(* IEC 61131-3 sources: SortJet_MasterSPS_Aufbau.fbsproj/09_Station/Stationen/_Basic, 3 files *)

(* ---- Basic_Glastransport_FB_V01_00_00.fb.st ---- *)
(* METADATA
{
	"v3Meta": {
		"objectGuid": "8cc859a4-3853-4716-ad69-f1a04cff8809"
	}
}
*)
FUNCTION_BLOCK Basic_Glastransport_FB_V01_00_00
VAR_INPUT

  // BOOL
  bpAktivieren                     : BOOL;
  bpEintransport                   : BOOL;
  bpEintransportRueckwaertig       : BOOL;
  bpAustransport                   : BOOL;
  bpAustransportRueckwaertig       : BOOL;
  bpVortransport                   : BOOL;
  bpVortransportRueckwaertig       : BOOL;
  bpMesskopplung                   : BOOL;
  bpDurchtransport                 : BOOL;
  bpGlaslaengenmessung             : BOOL;
  bpHandfahrenPlus                 : BOOL;
  bpHandfahrenMinus                : BOOL;
  bpScheibeZurueckFahren           : BOOL;
  bpScheibeVorFahren               : BOOL;
  bpAnforderungHandfunktion        : BOOL; // Handfunktionen greifen auch im Automatikbetrieb (z.B. waehrend der Bediener anlegt)
  bpScheibeQuittiert               : BOOL; // Bediener hat die Scheibe quittiert (Fehlmessung / Messergebnis)
  bpScheibeFreigegeben             : BOOL; // Scheibe ist nach der Messung freigegeben
  bpReferenz                       : BOOL;
  bpCheck                          : BOOL;
  bpReset                          : BOOL;
  bpAutomatikAktiv                 : BOOL;
  bpFreigabe                       : BOOL;
  bpMessrichtungNegativ            : BOOL;
  bpCheckMitVorgaenger             : BOOL;
  bpCheckMitNachfolger             : BOOL;
  bpRueckwaertigerTransport        : BOOL;
  bpScheibentrennen                : BOOL;
  bpAbbruchVortransport            : BOOL;

  // Sensoren
  bpSensorEinlauf                  : BOOL;
  bpSensorEinlaufVorAb             : BOOL;
  bpSensorAuslaufVorAb             : BOOL;
  bpSensorAuslauf                  : BOOL;

  // OPTIONEN
  bpOptionMessungSystemCheckAktiv            : BOOL;
  bpOptionMasterSlaveTransport               : BOOL;
  bpOptionScheibenmessungEintransport        : BOOL;
  bpOptionAustransportISOLinie               : BOOL;
  bpOptionSlaveAntrieb                       : BOOL;
  bpOptionNachSystemcheckAufAuslaufsensor    : BOOL;
  bpOptionbScheibenmessungSensorVorabAuslauf : BOOL;

  // WORD
  wlIndex : WORD := 0;

  // ENUM
  eGlastyp : GlasTyp_EN;

  // STRUCT
  InGlasTransportVorgaenger   : Interface_GlasTransport; // STRUKTUR: Informationen ueber den Aus- Ein- Transport der Vorgaengerstation
  InGlasTransportNachfolger   : Interface_GlasTransport; // STRUKTUR: Informationen ueber den Aus- Ein- Transport der Nachfolge- Station
  pAuftrag                    : Auftragsdaten_ST;            // AUFTRAG: Aktuelle daten zum Auftrag [Laenge, Hoehe, Modelle]
  stStationsNummern           : Station_ST;

  // POINTER
  ppParameterBaustein          : REFERENCE TO Parameter_Glastransport;
  ppAntriebsInformationen      : REFERENCE TO AntriebsInformationen;
  ppAntriebsInformationenSlave : REFERENCE TO AntriebsInformationen; // Wird nur verwendet um die Box Nummer anzeigen zu lassen

  // Antrieb
  Antrieb       : REFERENCE TO Rexroth_ctrlX_Drive_Eckelmann_MC_V01_02_02;
  Antrieb_Slave : REFERENCE TO Rexroth_ctrlX_Drive_Eckelmann_MC_V01_02_02;

END_VAR

VAR_OUTPUT

  // BOOL
  bpDone                        : BOOL;
  bpFehler                      : BOOL;
  bprtScheibe                   : BOOL; // Scheibenzaehler: Bool der wie ein Trigger genutzt wird
  bpStationBelegt               : BOOL;
  bpVerfahrFreigabe             : BOOL;
  bpScheibeFaehrtUeberAuslauf   : BOOL; // HINWEIS: Glas ist ueber den Auslauf-Sensor gefahren und somit in den Verfahrbereich des Transportshuttles -> Nehmen der Verfahrfreigabe fuer das Transportshuttles
  bpScheibeFaehrtUeberEinlauf   : BOOL;
  bpResetAbgeschlossen          : BOOL; // STATUS: Reset wurde abgeschlossen TRUE / FALSE
  bpOutBereitZumAustransport    : BOOL; // OUT STATUS: Bereit zum Austransport [Eintransport auf die Nachfolgerstation]
  bpAnforderungMessergebnis     : BOOL; // STATUS: Riemen wartet auf das Scann- Ergebnis aus dem Uebergeordneteten Baustein
  bpOutBereitZumEintransport    : BOOL; // OUT STATUS: Bereit zum Eintransport [Austransport auf die Vorgaengerstation]
  bpFreigabeFremdprozess        : BOOL;
  bpSlaveAktiv                  : BOOL;
  bpDurchtransportWarAktiv      : BOOL;
  bpUebergrosseScheibeUebergang : BOOL;

  // WORD
  wpFehlerNr                   : Fehlerkonstanten_EN;

  // DWORD
  dwpWartezeit                 : DWORD; // STATISTIK: Zeitwerte fuer die Statistik zum auswerten

  // REAL
  rpOutGeschwindigkeit         : REAL;
  rpGemesseneGlaslaenge        : REAL;

END_VAR

VAR

  // HARDWARE EINGAENGE (vom Umrichter)
  in_bSensorEinlauf             : BOOL;
  in_bSensorEinlaufVorAb        : BOOL;
  in_bSensorAuslaufVorab        : BOOL;
  in_bSensorAuslauf             : BOOL;

  // BOOL
  blErsterZyklus                : BOOL := TRUE;
  blScheibenMerker              : BOOL;
  blReduzierteGeschwindigkeit   : BOOL;
  blAntriebsKopplungAktiv       : BOOL;
  blStarteSlaveKopplung         : BOOL;
  blSlaveKopplungHergestellt    : BOOL; // Kopplung in dieser Anforderung neu hergestellt (SYNC_AUF_MASTER fertig)

  // INT
  ilScheibenZaehler             : INT;
  ilIndexScheibenmessung        : INT := 1;

  // REAL
  rlGefahreneStreckeEintransport    : REAL; // HINWEIS: Weg-Merker fuer die Strecke die beim Eintransport zurueck gelegt werden muss laut Auftrag
  rlPositionAntriebBeiStart         : REAL;
  rlMaxStreckeErsteScheibe          : REAL; // Max. Weg bis zur ersten Scheibe: Laenge der abgebenden Station, ohne bekannte Laenge die eigene Stationslaenge
  rlGlasgewicht                     : REAL;
  rlPositionScheibenAnfangErkannt   : REAL;
  rlStreckeBisZurVerzoegerung       : REAL;
  rlScheibenMessung                 : ARRAY[1..10] OF REAL;

  // STEPS
  steplEintransport             : Steps_TE;
  steplEintransportRueckwaertig : Steps_TE;
  steplAustransport             : Steps_TE;
  steplAustransportRueckwaertig : Steps_TE;
  steplVortransport             : Steps_TE;
  steplVortransportRueckwaertig : Steps_TE;
  steplDurchtransport           : Steps_TE;
  steplMesskopplung             : Steps_TE;
  steplGlaslaengenMessung       : Steps_TE;
  steplCheck                    : Steps_TE;
  steplReset                    : Steps_TE;
  steplReferenz                 : Steps_TE;
  steplSlave                    : Steps_TE;

  // TIMER
  toflAutoAbschaltung                       : TOF;
  toflEinlaufsensor                         : TOF;
  toflAuslaufsensor                         : TOF;
  tonlEinlaufsensor                         : TON; // Entprellung belegt (Flackern quittiert keine zweite Scheibe)
  tonlAuslaufsensor                         : TON; // Entprellung belegt (Flackern quittiert keine zweite Scheibe)
  toflVorAbStopSensorAuslauf                : TOF;
  toflVorAbStopSensorEinlauf                : TOF;
  tonlMaximaleZeitAuslaufsensorFreiFahren   : TON;
  tonlMaximaleZeitEinlaufsensorFreiFahren   : TON;
  tonlMaximaleZeitSensorAnfahren            : TON;
  tonlMaxWarteAufResetErfolgreich           : TON;
  tonlMaxWartezeitFremdanlage               : TON;
  tonlAntriebNichtBetriebsBereit            : TON;
  tonlSchrittueberwachung                   : TON;
  tonlUberwachungSlaveAktiv                 : TON;
  tonlSlaveKopplungDeaktiviert              : ton;
  tonlSlaveKopplungHerstellen               : TON; // Ueberwachung: Kopplung nicht hergestellt

  rtlMessungOK                              : R_TRIG;

  // TIME
  tlWarteZeitAufnahme    : TIME; // STATISTIK

  // TRIGGER
  ftlScheibeZurueckFahren : F_TRIG;
END_VAR

VAR_INPUT

  // BAUSTEINE
  Scheibenmessung  : Scheibenmessung_FB_V01_00_00;

END_VAR

VAR CONSTANT

  // TIME
  cUEBERWACHUNG_SLAVE_AKTIV           : TIME := T#1S;
  cMAX_ZEIT_SLAVE_KOPPLUNG_HERSTELLEN : TIME := T#30S; // inkl. Referenzfahrt von Master und Slave

END_VAR

//-------------------------------------------------------------------------------------------------
// INITIALISIERUNG
//-------------------------------------------------------------------------------------------------
IF ( blErsterZyklus ) THEN

  IF ( __ISVALIDREF(ppAntriebsInformationen) ) THEN

    blErsterZyklus            := FALSE;

    // Antrieb referenzieren
    Antrieb       REF= pgAntriebe[ppAntriebsInformationen.wAchsID];
    IF ( __ISVALIDREF(ppAntriebsInformationenSlave) ) THEN
      Antrieb_Slave REF= pgAntriebe[ppAntriebsInformationenSlave.wAchsID];
    END_IF

    (* Hinweis:
       - Initialisierung Antriebsinformationen
    *)
    Antrieb.ppAntriebsInformationen REF= ppAntriebsInformationen;
    Antrieb.stStationsNummern := stStationsNummern;
    IF ( __ISVALIDREF(Antrieb_Slave) AND __ISVALIDREF(ppAntriebsInformationenSlave) ) THEN
      Antrieb_Slave.ppAntriebsInformationen REF= ppAntriebsInformationenSlave;
      Antrieb_Slave.stStationsNummern := stStationsNummern;
    END_IF

    (* Hinweis:
       - Für die Zielpunktkontrolle muss im ersten Zyklus die Zielposition initialisiert werden
    *)
    Antrieb.rpZielPosition := Antrieb.rpIstPosition;
    IF ( __ISVALIDREF(Antrieb_Slave) AND __ISVALIDREF(ppAntriebsInformationenSlave) ) THEN
      Antrieb_Slave.rpZielPosition := Antrieb_Slave.rpIstPosition;
    END_IF

    (* Hinweis:
       - Antriebswerte vorinitialisieren
    *)
    Antrieb.rpGeschwindigkeit := ppAntriebsInformationen.rpMaxGeschwindigkeit;
    Antrieb.rpBeschleunigung  := ppAntriebsInformationen.rpMaxBeschleunigung;
    Antrieb.rpVerzoegerung    := ppAntriebsInformationen.rpMaxVerzoegerung;
    Antrieb.rpRuckzeit        := ppAntriebsInformationen.rpMaxRuckzeit;

    (* Hinweis:
       - Antriebswerte vorinitialisieren
    *)
    IF ( __ISVALIDREF(Antrieb_Slave) AND __ISVALIDREF(ppAntriebsInformationenSlave) ) THEN
      Antrieb_Slave.rpGeschwindigkeit := REAL#0;
      Antrieb_Slave.rpBeschleunigung  := ppAntriebsInformationenSlave.rpMaxBeschleunigung;
      Antrieb_Slave.rpVerzoegerung    := ppAntriebsInformationenSlave.rpMaxVerzoegerung;
      Antrieb_Slave.rpRuckzeit        := ppAntriebsInformationenSlave.rpMaxRuckzeit;
    END_IF

    // Pointer
    //   - Initialisierung zur vermeidung von null Pointerexceptions
    //     => Scheibenmessung
    Scheibenmessung.ppAntriebsInformationen REF= ppAntriebsInformationen;
    Scheibenmessung.ppAntrieb               REF= Antrieb;
    Scheibenmessung.pbpVorstopSensor        REF= bgFALSE;
    Scheibenmessung.pbpEinlaufSensor        REF= bgFALSE;

  ELSE
    RETURN;
  END_IF

END_IF

//-------------------------------------------------------------------------------------------------
// DEAKTIVIEREN
//-------------------------------------------------------------------------------------------------
IF ( NOT bpAktivieren ) THEN

  bpVerfahrFreigabe := TRUE;
  bpDone := TRUE;

  (* Hinweis:
     - Ausnahmesituationen
  *)
  bpFehler   := FALSE;
  wpFehlerNr := cMELDUNG_NULL;

  RETURN;

END_IF

//-------------------------------------------------------------------------------------------------
// IO ZUWEISUNG
//-------------------------------------------------------------------------------------------------
in_bSensorEinlauf      := Antrieb.udipEingaengeUmrichter.cXG31_1_I_1;
in_bSensorEinlaufVorAb := Antrieb.udipEingaengeUmrichter.cXG31_6_I_4;
in_bSensorAuslaufVorab := Antrieb.udipEingaengeUmrichter.cXG31_7_I_5;
in_bSensorAuslauf      := Antrieb.udipEingaengeUmrichter.cXG31_2_I_2;

bpSensorEinlauf      := in_bSensorEinlauf;
bpSensorEinlaufVorAb := in_bSensorEinlaufVorAb;
bpSensorAuslaufVorab := in_bSensorAuslaufVorab;
bpSensorAuslauf      := in_bSensorAuslauf;

//-------------------------------------------------------------------------------------------------
// TIMER, SETTINGS, ETC.
//-------------------------------------------------------------------------------------------------
// Sensorenflackern
toflEinlaufsensor(IN := bpSensorEinlauf, PT := T#50MS);
toflAuslaufsensor(IN := bpSensorAuslauf, PT := T#50MS);
tonlEinlaufsensor(IN := bpSensorEinlauf, PT := T#50MS);
tonlAuslaufsensor(IN := bpSensorAuslauf, PT := T#50MS);
toflVorAbStopSensorEinlauf(IN := bpSensorEinlaufVorab, PT := t#50ms);
toflVorAbStopSensorAuslauf(IN := bpSensorAuslaufVorAb, PT := t#50ms);

// Reset
tonlMaxWarteAufResetErfolgreich(IN:=bpReset,pt:=tgMaxWartezeitReset-T#1S);

//-------------------------------------------------------------------------------------------------
// AUFRUFE
//-------------------------------------------------------------------------------------------------
// 2. Riemen/Rollen vorhanden -> Kipptisch
//   - Vor den Schrittketten, damit diese die Kopplung im selben Zyklus sehen
//   - Kopplung gilt, wenn der Slave synchron ist, die Kopplung angefordert ist und in dieser Anforderung
//     neu hergestellt wurde (sonst gilt beim direkten Wechsel z. B. Eintransport -> Vortransport noch kurz
//     das alte Synchron-Signal des Antriebs, und die neue Kette meldet "Slave-Kopplung verloren")
IF bpOptionSlaveAntrieb THEN
  SlaveAntrieb();
  blAntriebsKopplungAktiv := Antrieb_Slave.bpAchseSychron AND blStarteSlaveKopplung AND blSlaveKopplungHergestellt;
ELSE
  blAntriebsKopplungAktiv := TRUE;
END_IF

Eintransport();
Eintransport_Rueckwaertig();
Vortransport();
Vortransport_Rueck();
Durchtransport();
Messkopplung();
Laengenmessung();
SystemCheck();
Referenz();
Handfunktionen();
Meldungen();
Reset();

IF ( bpOptionAustransportISOLinie ) THEN
  Austransport_ISO();
  Austransport_Rueckwaertig_ISO();
ELSIF ( bpOptionMasterSlaveTransport ) THEN
  Austransport_MasterSlave();
  Austransport_Rueckwaertig_MasterSlave();
ELSE
  Austransport();
  Austransport_Rueckwaertig();
END_IF

//-------------------------------------------------------------------------------------------------
// FREIGABEN UND AUFRUFE
//-------------------------------------------------------------------------------------------------
// Glastransportfreigabe
//   - Freigabe
toflAutoAbschaltung( IN := (  bpAutomatikAktiv
                             AND ( bpAustransport
                                   OR bpAustransportRueckwaertig
                                   OR bpEintransport
                                   OR bpEintransportRueckwaertig
                                   OR bpVortransport
                                   OR bpVortransportRueckwaertig
                                   OR bpMesskopplung
                                   OR bpDurchtransport
                                   OR bpGlaslaengenmessung
                                 ) )
                     OR bpCheck
                     OR bpHandfahrenMinus
                     OR bpHandfahrenPlus
                     OR bpScheibeZurueckFahren
                     OR bpReferenz,
                     PT:= tgZeitAutoabschaltungEnergiesparModus );

// Aufruf:
//   - Antriebe
//   - Scheibenmessung
Antrieb.bpFreigabe        := toflAutoAbschaltung.Q AND bpFreigabe;
Antrieb.rpRuckzeit        := ppAntriebsInformationen.rpMaxRuckzeit;
Antrieb.stStationsNummern := stStationsNummern;

IF bpOptionSlaveAntrieb THEN
  Antrieb_Slave.bpFreigabe        := Antrieb.bpFreigabe;
  Antrieb_Slave.rpRuckzeit        := ppAntriebsInformationen.rpMaxRuckzeit;
  Antrieb_Slave.stStationsNummern := stStationsNummern;
END_IF

Scheibenmessung( stStationsNummern                   := stStationsNummern,
                 ppAntrieb                           := Antrieb,
                 pbpVorstopSensor                    := bpSensorAuslaufVorab,
                 pbpEinlaufSensor                    := bpSensorEinlauf,
                 bpDrehrichtungsumkehrMessung        := bpMessrichtungNegativ,
                 rpMessstrecke                       := ppParameterBaustein.rMessstrecke,
                 ppAntriebsInformationen             := ppAntriebsInformationen,
                 bpAuswahlSensorVorabScheibenmessung := bpOptionbScheibenmessungSensorVorabAuslauf,
                 rpFaktorBremswegverlaengern         := 1.6 ) ;

//-------------------------------------------------------------------------------------------------
// AKTION AUSGAENGE
//-------------------------------------------------------------------------------------------------
// Ausgaeng:
//   - Aktuelle Geschwindigkeit des Antriebs
//     -> Soll- Wertkopplung ( Soll-Geschwindigkeit des Antriebs)
//     -> Ist- Wertkopplung ( Soll-Geschwindigkeit des Antriebs)
IF ( ( bpEintransport OR bpEintransportRueckwaertig ) AND bpOutBereitZumEintransport )THEN
  rpOutGeschwindigkeit :=  ABS(Antrieb.rpGeschwindigkeit);
ELSE
  rpOutGeschwindigkeit :=  ABS(Antrieb.rpIstGeschwindigkeit);
END_IF

// Freigabe für eine Bewegung
bpVerfahrFreigabe :=  NOT ( bpSensorEinlauf
                            OR bpSensorAuslauf
                            OR bpEintransport
                            OR bpAustransport );
END_FUNCTION_BLOCK

(* ---- Basic_Schnittstelle_FB_V01_00_00.fb.st ---- *)
(* METADATA
{
	"v3Meta": {
		"objectGuid": "466fafaa-eb0c-4cc2-9ac3-d488ea338d40"
	}
}
*)
FUNCTION_BLOCK Basic_Schnittstelle_FB_V01_00_00
VAR_IN_OUT

  // STRUKT
  BasisStationsParameter     : StationBasisParameter_ST;

END_VAR

VAR_INPUT

  // BOOL
  bpEmpfaengerSensorEinlauf  : BOOL;
  bpResetISOLinieEvent       : BOOL;
  bpStarteIGEvent            : BOOL;

  // WORD
  wpAuftragsTyp              : WORD; // Unterteilung => 0 = Scheibe vom Sortjet , 1 = Scheibe soll Manuell angelegt werden *)

  // STRUCT
  AuftragsSpeicher           : Auftragswarteschlange_Fremdanlage_FB;

END_VAR

VAR_OUTPUT

  // BOOL
  bpISOLineEventAktiv       : BOOL; // Offenes ISO Linie Event nach aussen weitergeben

  // REAL
  rpGeschwindigkeit          : REAL;

  //DWORD
  dwpWartezeit     : DWORD;// STATISTIK: Beschreibt die Zeit zwischen Anlegeauftrag und betaetigen des Tasters zum Eintransport

END_VAR

VAR

  // BOOL
  blErsterZyklus             : BOOL := TRUE;
  bEmpfaengerSensorEinlauf   : BOOL; // Eingang Einlaufsensor von Umrichter Box
  blBereitZumEintransport    : BOOL;
  blBereitZumAustransport    : BOOL;
  blAutomatikBetriebAktiv    : BOOL;
  blSenderBereit             : BOOL;
  blSenderGlasBereit         : BOOL;
  blInLogSchreiben           : BOOL;
  blOutLogSchreiben          : BOOL;
  blTempSenderBereit         : BOOL;
  blTempSenderGlasBereit     : BOOL;
  blTempFreigabeSK           : BOOL;
  blTempAnforderungSK        : BOOL;
  blTempGlasAbruf            : BOOL;
  blTempEinlaufSensor        : BOOL;
  blTempAutomatikBetrieb     : BOOL;
  blUebergabeGlas            : BOOL; // Schrittkettenvariable
  blStartISOLinie            : BOOL; // Schrittkettenvariable

  // WORD
  wlWatchIONachrichtenNummer : WORD;

  //TRIGGER
  rtlTasterSpezial           : R_TRIG;
  rtlTasterGlasbruch         : R_TRIG;

  // STRING
  slInLogString              : STRING;
  slOutLogString             : STRING;

  // TIME
  tlWarteZeiteAufnahme       : TIME;

  // STEPS
  steplUebergabeGlas         : Steps_TE;

  // BAUSTEINE
  Horn                       : Horn_FB;

  // GLAETTUNG AUSGANGSGESCHWINDIGKEIT (M_GeschwindigkeitGlaetten)
  blGeschwindigkeitInitialisiert     : BOOL; // Erste Geschwindigkeit nach Stillstand uebernommen
  blGeschwindigkeitUpdateSperreAktiv : BOOL; // Sperrzeit nach Geschwindigkeitsaenderung aktiv
  rlGeschwindigkeitFreigegeben       : REAL; // Zuletzt freigegebene Geschwindigkeit
  tonlGeschwindigkeitUpdateSperre    : TON;

END_VAR

VAR_INPUT

  // HARDWARE EINGAENGE
  in_bEmpfaengerSensorEinlauf         : BOOL; // Einlaufsensor
  in_bTasterGlasbruch           AT%I* : BOOL; // Taster, Gegenscheibe wurde ausgeschleust
  in_bTasterSpezial             AT%I* : BOOL; // Taster, Sonderscheibe zugestellt

  // HARDWARE AUSGAENGE
  out_bSenderBereit             AT %Q* : BOOL; // Anlage zum Transport bereit
  out_bSenderGlasBereit         AT %Q* : BOOL; // Glas bereit zum Transport
  out_bLeuchteGlasbruch         AT %Q* : BOOL;
  out_bLeuchteSpezial           AT %Q* : BOOL;
  out_bAmpelEventAktiv          AT %Q* : BOOL;

END_VAR

//-------------------------------------------------------------------------------------------------
// INITIALISIERUNG
//-------------------------------------------------------------------------------------------------
IF ( blErsterZyklus ) THEN
  blErsterZyklus:=FALSE;

END_IF

//-------------------------------------------------------------------------------------------------
// BAUSTEIN: DEAKTIVIERUNG
//-------------------------------------------------------------------------------------------------
(* Hinweis:
   - Schnittstelle deaktiviert (MK bDeaktivieren): Ausgaenge zur Fremdanlage abschalten, Baustein verlassen.
     Abgeleitete Bausteine pruefen nach SUPER^() selbst und schalten ihre eigenen Ausgaenge ab
*)
IF ( BasisStationsParameter.stMKs.bDeaktivieren ) THEN
  out_bSenderBereit     := FALSE;
  out_bSenderGlasBereit := FALSE;
  out_bLeuchteGlasbruch := FALSE;
  out_bLeuchteSpezial   := FALSE;
  out_bAmpelEventAktiv  := FALSE;
  bpISOLineEventAktiv   := FALSE;
  rpGeschwindigkeit     := 0;
  RETURN;
END_IF

//-------------------------------------------------------------------------------------------------
// AKTIONEN
//-------------------------------------------------------------------------------------------------
IF ( BasisStationsParameter.bReset ) THEN
  Reset();
END_IF

IF ( BasisStationsParameter.stMKs.stFremdanlage.bAnzeigeISOLinieEventAktiv ) THEN
  IGLineEvent();
END_IF

A_Schnittstelle();

//-------------------------------------------------------------------------------------------------
// BAUSTEIN: ZUWEISUNGEN, AUFRUFE
//-------------------------------------------------------------------------------------------------
Horn(bpAktiv := bgHornAktivieren);
END_FUNCTION_BLOCK

(* ---- Basic_Station_FB_V01_00_00.fb.st ---- *)
(* METADATA
{
	"v3Meta": {
		"objectGuid": "b8afb014-b2bc-4dd4-b6e0-59869c47ec49"
	}
}
*)
FUNCTION_BLOCK Basic_Station_FB_V01_00_00
VAR_IN_OUT

  // STRUKT
  BasisStationsParameter : StationBasisParameter_ST;

END_VAR

VAR_INPUT

END_VAR

VAR_OUTPUT

  // DWORD
  dwpHandfunktionenReturn    : DWORD; // Aktive Handfunktionen, gleiche Bitbelegung wie dwlHandfunktionen (Aktion HandfunktionenStatus der Station)

END_VAR

VAR

  // BOOLEAN
  blErsterZyklus             : BOOL := TRUE; // Initialisierung
  blBetriebsartHand          : BOOL;
  blBetriebsartReset         : BOOL;
  blBetriebartCheck          : BOOL;
  blBetriebsartAutomatik     : BOOL;
  blBetriebsartReferenz      : BOOL;
  blMerkerFehlerAutomatik    : BOOL;
  blNachSystemcheckMerker    : BOOL; // Merkt sich, wenn der Systemcheck erfolgreich durchgeführt wurde, damit die Gebläse nicht nach dem Systemcheck ausgehen

  // WORD
  wlBetriebsart              : WORD;
  wlWatchIONachrichtenNummer : WORD;
  wlIndex                    : WORD;

  // DWORD
  dwlHandfunktionen                : DWORD;  // Handfunktionen: 0..31 Bit
  dwlHandfunktionenZuletztGesendet : DWORD;  // Rueckmeldung der Handfunktionen zum MMI

  // STEPS
  steplReset                 : Steps_TE;
  steplCheck                 : Steps_TE;
  steplReferenz              : Steps_TE;
  steplEintransport          : Steps_TE;
  steplAustransport          : Steps_TE;
  steplVortransport          : Steps_TE;
  steplDurchtransport        : Steps_TE;
  steplMesskopplung          : Steps_TE;
  steplAnlegen               : Steps_TE;
  steplAbnehmen              : Steps_TE;
  steplGlaslaengenmessung    : Steps_TE;
  steplGlashoehenmessung     : Steps_TE;
  steplPositionieren         : Steps_TE;

  // TRIGGER
  ftlBausteinDeaktivierung              : F_TRIG;
  rtlFehlerMeldungGenerierenHandbetrieb : R_TRIG;

  // TIMER
  tonlMaxWarteAufResetErfolgreich       : TON;

END_VAR

//-------------------------------------------------------------------------------------------------
// INITIALISIERUNG UND EINSTELLUNGEN
//-------------------------------------------------------------------------------------------------
IF ( blErsterZyklus  ) THEN

  blErsterZyklus := FALSE;

  // Initialisierung des Bausteins
  A_Baustein_Initialisierung();

END_IF

//-------------------------------------------------------------------------------------------------
// DEAKTIVIERUNG DES BAUSTEINS
//-------------------------------------------------------------------------------------------------

// Werte wieder passend abloeschen, wenn der Baustein wieder aktiviert wird
ftlBausteinDeaktivierung( CLK := BasisStationsParameter.stMKs.bDeaktivieren );

IF ( ftlBausteinDeaktivierung.Q ) THEN

  FOR wlIndex := cWAND_1 TO cANZAHL_WAENDE DO
    BasisStationsParameter.bAustransportAbgeschlossen[wlIndex]   := FALSE;
    BasisStationsParameter.bDurchtransportAbgeschlossen[wlIndex] := FALSE;
    BasisStationsParameter.bEintransportAbgeschlossen[wlIndex]   := FALSE;
    BasisStationsParameter.bMesskopplungAbgeschlossen[wlIndex]   := FALSE;
    BasisStationsParameter.bVorabKomponentenAnsteuerungAbgeschlossen[wlIndex] := FALSE;
    BasisStationsParameter.bVortransportAbgeschlossen[wlIndex]   := FALSE;
    BasisStationsParameter.bStationBelegt[wlIndex]               := FALSE;
  END_FOR

  BasisStationsParameter.bFehler                := FALSE;
  BasisStationsParameter.wFehlerNummer          := cMELDUNG_NULL;
  BasisStationsParameter.bAuftragAktiv          := FALSE;
  BasisStationsParameter.bReset                 := FALSE;
  BasisStationsParameter.bIstReferenziert       := FALSE;
  BasisStationsParameter.bCheckAbgeschlossen    := FALSE;
  BasisStationsParameter.bReferenzAbgeschlossen := FALSE;

END_IF

(* Hinweis:
   - Deaktivierung des Bausteins
     => Der Baustein wird zum Ende der RETURN-Anweisung verlassen
*)
IF ( BasisStationsParameter.stMKs.bDeaktivieren ) THEN

  A_ScheibenDeaktivierteStationMelden();

  FOR wlIndex := cWAND_1 TO cANZAHL_WAENDE DO
    BasisStationsParameter.bAustransportAbgeschlossen[wlIndex]   := TRUE;
    BasisStationsParameter.bDurchtransportAbgeschlossen[wlIndex] := TRUE;
    BasisStationsParameter.bEintransportAbgeschlossen[wlIndex]   := TRUE;
    BasisStationsParameter.bMesskopplungAbgeschlossen[wlIndex]   := TRUE;
    BasisStationsParameter.bVorabKomponentenAnsteuerungAbgeschlossen[wlIndex] := TRUE;
    BasisStationsParameter.bVortransportAbgeschlossen[wlIndex]   := TRUE;
    BasisStationsParameter.bStationBelegt[wlIndex]               := FALSE;
  END_FOR

  BasisStationsParameter.bAbnehmenAbgeschlossen := TRUE;
  BasisStationsParameter.bAnlegenAbgeschlossen := TRUE;
  BasisStationsParameter.bCheckAbgeschlossen    := TRUE;
  BasisStationsParameter.bGlashoehenmessungAbgeschlossen := TRUE;
  BasisStationsParameter.bGlaslaengenmessungAbgeschlossen := TRUE;
  BasisStationsParameter.bReferenzAbgeschlossen := TRUE;
  BasisStationsParameter.bVorabDrehenAbgeschlossen := TRUE;
  BasisStationsParameter.bVorabpositionierenAbgeschlossen := TRUE;
  BasisStationsParameter.bIstReferenziert       := TRUE;

  BasisStationsParameter.bReset        := FALSE;
  BasisStationsParameter.bFehler := FALSE;
  BasisStationsParameter.wFehlerNummer := cMELDUNG_NULL;
  BasisStationsParameter.bAuftragAktiv := FALSE;

  RETURN;

END_IF

//-------------------------------------------------------------------------------------------------
// AKTIONEN
//-------------------------------------------------------------------------------------------------
A_Schnittstelle();
Betriebsart();
Meldungen();

//-------------------------------------------------------------------------------------------------
// TIMER
//-------------------------------------------------------------------------------------------------
// Reset
tonlMaxWarteAufResetErfolgreich( IN := BasisStationsParameter.bReset, PT := tgMaxWartezeitReset);
END_FUNCTION_BLOCK
